KUKA KRL program: LongProg1.src

&ACCESS RVP
&REL 1
&PARAM TEMPLATE = C:\KRC\Roboter\Template\vorgabe
&PARAM EDITMASK = *
DEF LongProg1 ( )

; External program calls:
EXT LongProg2()

; ---- Setting tool (TCP) ----
$TOOL = {FRAME: X 10.000,Y 20.000,Z 150.000,A 0.000,B 0.000,C 0.000}
; --------------------------
PTP {A1 0.00000,A2 -10.00000,A3 20.00000,A4 0.00000,A5 30.00000,A6 0.00000}
PTP {A1 20.00000,A2 -10.00000,A3 20.00000,A4 0.00000,A5 30.00000,A6 0.00000}

; Continue running program as cascaded execution
LongProg2()

END
